Fanuc KAREL source: ko00070.KL

-- PROVISIONAL review KL for V770-1; original PC SHA256 80e86f9d99b508026d32a8b0efb1187ae14178167acf41ad3346a7e943211167
-- Incomplete behavior may be omitted. Consult companion uncertainty JSON. Do not deploy.
PROGRAM KO00070
%NOLOCKGROUP
BEGIN
  -- UNRESOLVED_PC offsets 5-12; opcodes 9D,23
  -- UNRESOLVED_PC offsets 17-66; opcodes 27,22,1C,27,49,7E,AD,22,31,7E,4A
  -- UNRESOLVED_PC offsets 71-75; opcodes 7F
END KO00070
